{attribute 'qualified_only'}
{attribute 'strict'}
{attribute 'to_string'}
TYPE E_TriBlenderUsage :
(
	eNotInUse := 0,
	eMarinada_T1,
	eMarinada_T2,
	eMarinada_Standby,
	eColor_T3,
	eColor_T4,
	eColor_Standby
);
END_TYPE

(* stored: Version 1.1.0.1, ProductVersion 3.1.4024.12
   DUT E_TriBlenderUsage: Id {a2f2d29e-a9a2-4788-996c-f36425cb4241} *)
